VAR_GLOBAL CONSTANT
	mF_Mpc_degrees: DINT := 3;
	mF_Mpc_voff: LREAL := 0.0;
	mF_Mpc_yoff: LREAL := 0.05;
	mF_Mpc_RYscale: LREAL := 1.0;
	mF_Mpc_RMDscale: LREAL := 1.0;
	mF_Mpc_myoff: LREAL := 0.05;
	SS_INITIALIZE: SINT := 0;
	SS_STEP: SINT := 1;
END_VAR

(* stored: Version 1.1.0.1, ProductVersion 3.1.4024.9
   GVL GVL_1664200802: Id {fdcf1e7e-0072-4c57-a086-f54a2cea0b67} *)
